ABB RAPID module: Module1_0915含四个练习.mod

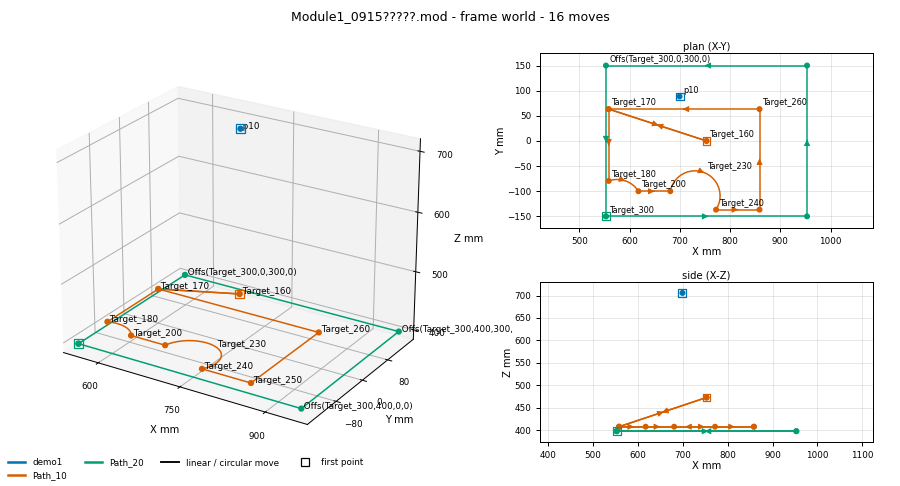
[picture p0: tool path of Module1_0915含四个练习.mod in frame world, 16 of 16 moves have a stored position in this frame; points joined in program order, loops and branches not executed]
MODULE Module1
    CONST robtarget p10:=[[699.42,88.43,705.75],[0.190432,-0.061687,0.979687,0.0119907],[0,0,0,0],[9E+9,9E+9,9E+9,9E+9,9E+9,9E+9]];
    CONST robtarget p20:=[[699.42,88.43,705.75],[0.190432,-0.061687,0.979687,0.0119907],[0,-1,0,0],[9E+9,9E+9,9E+9,9E+9,9E+9,9E+9]];
    CONST robtarget p30:=[[762.23,96.37,426.55],[0.00469136,-0.0628409,0.998012,0.000295343],[0,-1,0,0],[9E+9,9E+9,9E+9,9E+9,9E+9,9E+9]];
    CONST robtarget Target_160:=[[752.961021712,0,473.000001678],[-0.00000002,0,1,0],[0,-1,0,0],[9E+09,9E+09,9E+09,9E+09,9E+09,9E+09]];
    CONST robtarget Target_170:=[[558.409,63.326,408],[0,0,1,0],[0,-1,0,0],[9E+09,9E+09,9E+09,9E+09,9E+09,9E+09]];
    CONST robtarget Target_180:=[[558.409,-79.547,408],[0,0,1,0],[-1,0,-1,0],[9E+09,9E+09,9E+09,9E+09,9E+09,9E+09]];
    CONST robtarget Target_190:=[[591.551,-79.397,408],[0,0,1,0],[-1,0,-1,0],[9E+09,9E+09,9E+09,9E+09,9E+09,9E+09]];
    CONST robtarget Target_200:=[[617.506,-100.006,408],[0,0,1,0],[-1,0,-1,0],[9E+09,9E+09,9E+09,9E+09,9E+09,9E+09]];
    CONST robtarget Target_210:=[[752.961,0,473],[0,0,1,0],[0,0,0,0],[9E+09,9E+09,9E+09,9E+09,9E+09,9E+09]];
    CONST robtarget Target_220:=[[680.926,-100.006,408],[0,0,1,0],[0,0,0,0],[9E+09,9E+09,9E+09,9E+09,9E+09,9E+09]];
    CONST robtarget Target_230:=[[748.721,-63.019,408],[0,0,1,0],[0,0,0,0],[9E+09,9E+09,9E+09,9E+09,9E+09,9E+09]];
    CONST robtarget Target_240:=[[771.941,-136.674,408],[0,0,1,0],[0,0,0,0],[9E+09,9E+09,9E+09,9E+09,9E+09,9E+09]];
    CONST robtarget Target_250:=[[858.409,-136.674,408],[0,0,1,0],[0,0,0,0],[9E+09,9E+09,9E+09,9E+09,9E+09,9E+09]];
    CONST robtarget Target_260:=[[858.409,63.326,408],[0,0,1,0],[0,0,0,0],[9E+09,9E+09,9E+09,9E+09,9E+09,9E+09]];
    CONST robtarget Target_270:=[[558.409,63.326,408],[0,0,1,0],[0,0,0,0],[9E+09,9E+09,9E+09,9E+09,9E+09,9E+09]];
    CONST robtarget Target_280:=[[752.961,0,473],[0,0,1,0],[0,0,0,0],[9E+09,9E+09,9E+09,9E+09,9E+09,9E+09]];
    CONST robtarget Target_300:=[[552.961,-150,398],[-0.00000002,0,1,0],[0,0,0,0],[9E+09,9E+09,9E+09,9E+09,9E+09,9E+09]];
    CONST robtarget Target_310:=[[752.96,0.00,473.00],[4.57512E-9,0,-1,0],[0,0,0,0],[9E+9,9E+9,9E+9,9E+9,9E+9,9E+9]];

    PROC main()
        !writewhattogood?
    ENDPROC

    PROC demo1()
        MoveJ p10,v200,z20,MyTool;
    ENDPROC

    PROC Path_10()
        MoveJ Target_160,v50,z100,MyTool\WObj:=wobj0;
        MoveL Target_170,v50,z100,MyTool\WObj:=wobj0;
        MoveL Target_180,v50,z100,MyTool\WObj:=wobj0;
        MoveC Target_190,Target_200,v50,z100,MyTool\WObj:=wobj0;
        MoveL Target_220,v50,z100,MyTool\WObj:=wobj0;
        MoveC Target_230,Target_240,v50,z100,MyTool\WObj:=wobj0;
        MoveL Target_250,v50,z100,MyTool\WObj:=wobj0;
        MoveL Target_260,v50,z100,MyTool\WObj:=wobj0;
        MoveL Target_270,v50,z100,MyTool\WObj:=wobj0;
        MoveL Target_280,v50,z100,MyTool\WObj:=wobj0;
    ENDPROC

    PROC Path_20()
        MoveL Target_300,v50,z100,MyTool\WObj:=wobj0;
        MoveL Offs(Target_300,400,0,0),v50,z100,MyTool\WObj:=wobj0;
        MoveL Offs(Target_300,400,300,0),v50,z100,MyTool\WObj:=wobj0;
        MoveL Offs(Target_300,0,300,0),v50,z100,MyTool\WObj:=wobj0;
        MoveL Target_300,v50,z100,MyTool\WObj:=wobj0;
    ENDPROC

    PROC swap_num()
        VAR num num1;
        VAR num num2;
        VAR num temp;
        VAR num key;
        TPErase;
        TPReadNum num1,"First num1 ->";
        TPReadNum num2,"Second num2 ->";
        temp:=num1;
        num1:=num2;
        num2:=temp;
        TPWrite "num1:"\Num:=num1;
        TPWrite "num2:"\Num:=num2;
        TPReadFK key,"Swap done. Press OK to finish","","","","OK","";
    ENDPROC

    PROC min_of_three()
        VAR num num1;
        VAR num num2;
        VAR num num3;
        VAR num min1;
        ! ?????
        VAR num key;
        TPErase;
        TPReadNum num1,"First num ->";
        TPReadNum num2,"Second num ->";
        TPReadNum num3,"Third num ->";
        min1:=num1;
        ! ? ?????????
        IF num2<min1 THEN
            min1:=num2;
            ! ? ????????
        ENDIF
        IF num3<min1 THEN
            min1:=num3;
            ! ? ????????
        ENDIF
        TPWrite "min"\Num:=min1;
        ! ?????
        TPReadFK key,"Min found. Press OK to finish","","","","OK","";
    ENDPROC

    PROC time_period()
        VAR num timeval;
        ! input value
        VAR num key;
        TPErase;
        TPReadNum timeval,"time?";
        IF timeval>=0 AND timeval<=5 THEN
            TPWrite "dawn";
            ! 0-5
        ELSEIF timeval>=6 AND timeval<=11 THEN
            TPWrite "morning";
            ! 6-11
        ELSEIF timeval>=12 AND timeval<=17 THEN
            TPWrite "afternoon";
            ! 12-17
        ELSEIF timeval>=18 AND timeval<=23 THEN
            TPWrite "evening";
            ! 18-23
        ELSE
            TPWrite "NG";
            ! others
        ENDIF
        TPReadFK key,"Done. Press OK to finish","","","","OK","";
    ENDPROC

    PROC library_fee()
        VAR num booktype;
        ! 1=Normal  2=Popular  3=Reference
        VAR num days;
        VAR num freedays;
        ! free days of the chosen type
        VAR num rate;
        ! fee per extra day
        VAR num price;
        VAR num key;
        TPErase;
        ! --- Step 1: choose book type (keys 1..3 enabled) ---
        TPReadFK booktype,"Select book type","Normal","Popular","Reference","","";
        ! --- Step 2: decide free days and rate by type ---
        IF booktype=1 THEN
            freedays:=14;
            rate:=0.5;
        ELSEIF booktype=2 THEN
            freedays:=7;
            rate:=0.8;
        ELSEIF booktype=3 THEN
            freedays:=3;
            rate:=1.2;
        ELSE
            freedays:=0;
            rate:=0;
        ENDIF
        ! --- Step 3: input days ---
        TPReadNum days,"Days?";
        ! --- Step 4: calculate the fee ---
        IF days>freedays THEN
            price:=(days-freedays)*rate;
        ELSE
            price:=0;
            ! within free days -> no fee
        ENDIF
        ! --- Step 5: show the result ---
        TPWrite "Price:"\Num:=price;
        TPReadFK key,"Done. Press OK to finish","","","","OK","";
    ENDPROC
ENDMODULE
